TYPE "ST_ConfigRecord"
VERSION : 0.1
   STRUCT
      Scope : String[80];
      WriteKey : String[160];
      Revision : UDInt;
      Kind : DInt;
      ValueType : DInt;
      ValueText : String[80];
   END_STRUCT;

END_TYPE

